Fanuc KAREL source: KT00427.KL

PROGRAM KT00427
%NOLOCKGROUP
VAR
  P1: XYZWPREXT
  P2: POSITION
  OUT: BOOLEAN
BEGIN
  P1.X = 1.0
  OUT = P1 > P2
END KT00427
